Staubli VAL3: saveCall.pgx

program saveCall()
begin
  if taskStatus("Save")==-1
    taskCreate "Save",100,saveTask()
  endIf
end
